(* Logix 5000 project; controller WWTP_CLX vendor 1 type 14 code 54 rev 17.2; software revision 17.00; part 12 of 13 *)
(* tags used below, declared in another part *)
   I_FeedP2_Fault : ALIAS FOR WWTP_CLX_Rack01_Slot00_CNB:I.Slot[1].Data.6;
   I_FeedP2_Fault_IOFault : ALIAS FOR WWTP_CLX_Rack01_Slot00_CNB:I.Slot[1].Fault.6;
   I_FeedP2_InAuto : ALIAS FOR WWTP_CLX_Rack01_Slot00_CNB:I.Slot[1].Data.4;
   I_FeedP2_InAuto_IOFault : ALIAS FOR WWTP_CLX_Rack01_Slot00_CNB:I.Slot[1].Fault.4;
   I_FeedP2_OverLoad : ALIAS FOR WWTP_CLX_Rack01_Slot00_CNB:I.Slot[1].Data.7;
   I_FeedP2_OverLoad_IOFault : ALIAS FOR WWTP_CLX_Rack01_Slot00_CNB:I.Slot[1].Fault.7;
   I_FeedP2_RunFdbk : ALIAS FOR WWTP_CLX_Rack01_Slot00_CNB:I.Slot[1].Data.5;
   I_FeedP2_RunFdbk_IOFault : ALIAS FOR WWTP_CLX_Rack01_Slot00_CNB:I.Slot[1].Fault.5;
   I_FeedP2_SpeedFdbk : ALIAS FOR WWTP_CLX_Rack01_Slot00_CNB:4:I.Ch3Data;
   I_FeedP2_SpeedFdbk_IOFault : ALIAS FOR WWTP_CLX_Rack01_Slot00_CNB:4:I.Ch3Fault;
   O_FeedP2_Out_Run : ALIAS FOR WWTP_CLX_Rack01_Slot00_CNB:2:O.Data.1;
   O_FeedP2_SpeedRef : ALIAS FOR WWTP_CLX_Rack01_Slot00_CNB:6:O.Ch1Data;
   O_FeedP2_SpeedRef_IOFault : ALIAS FOR WWTP_CLX_Rack01_Slot00_CNB:6:I.Ch1Fault;
   PLC_Device_ResetPB : BOOL;   // Site Wide Device Reset Push Button
   PLC_Simulation : BOOL;   // Application running IN SIMULATION
   WWTP_AerTk_InflFlow : UD_Flow;   // Aeration Tank Influent Flow
   WWTP_Alum : UD_Chemical;   // Alum Chemical
   WWTP_AlumTk1Lv : P_AIn;   // Alum Tank #1 Level
   WWTP_FeedP1 : UD_VSD;   // Feed Pump #1
   WWTP_FeedP1_FlowPacing : U_FlowPacing;   // Feed Pump #1 Flow Pacing
   WWTP_FeedP2 : UD_VSD;   // Feed Pump #2
   WWTP_FeedP2_FlowPacing : U_FlowPacing;   // Feed Pump #2 Flow Pacing
   WWTP_FeedP2_OverLoad : P_DIn;   // Feed Pump #2 Overload
   WWTP_FeedSys_OSet_PumpSelect : BOOL;   // Feed Pump System Pump Select
(* FeedP1, continued *)

ROUTINE Main   (* ladder *)
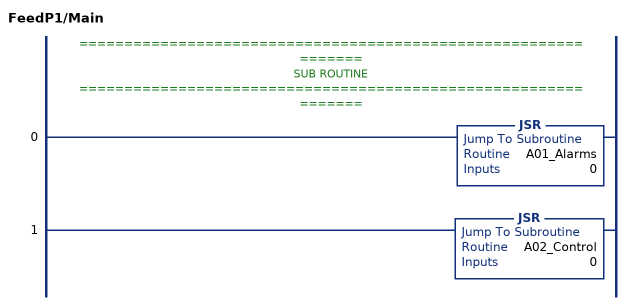
   // ===============================================================
   // SUB ROUTINE
   // ===============================================================
   0: JSR(A01_Alarms,0);
   1: JSR(A02_Control,0);
END_ROUTINE
END_PROGRAM

PROGRAM FeedP2   (* main routine Main *)
VAR
   Device : ALIAS FOR WWTP_FeedP2;
   Device_Alm0 : ALIAS FOR WWTP_FeedP2_OverLoad;
   Device_Alm0_Input : ALIAS FOR I_FeedP2_OverLoad;
   Device_Alm0_Input_IOFault : ALIAS FOR I_FeedP2_OverLoad_IOFault;
   Device_Alm1 : P_DIn := (Inp_Gate := 1, Cfg_NormTextVis := 1, Cfg_PCmdClear := 1, Cfg_TgtDisagreeAckReqd := 1, Cfg_TgtDisagreeSeverity := 3, Sts_InpPV := 1, Ack_TgtDisagree := 1, Rdy_SubstPV := 1);
   Device_Alm1_Input : BOOL;
   Device_Alm1_Input_IOFault : BOOL;
   Device_Alm2 : P_DIn := (Inp_Target := 1, Inp_Gate := 1, Cfg_NormTextVis := 1, Cfg_PCmdClear := 1, Cfg_TgtDisagreeAckReqd := 1, Cfg_TgtDisagreeSeverity := 3, Sts_SubstPV := 1, Sts_TgtDisagree := 1, Ack_TgtDisagree := 1, Rdy_InpPV := 1);
   Device_Alm2_Input : BOOL;
   Device_Alm2_Input_IOFault : BOOL;
   Device_Alm3 : P_DIn := (Inp_Target := 1, Inp_Gate := 1, Cfg_NormTextVis := 1, Cfg_PCmdClear := 1, Cfg_TgtDisagreeAckReqd := 1, Cfg_TgtDisagreeSeverity := 3, Sts_SubstPV := 1, Sts_TgtDisagree := 1, Ack_TgtDisagree := 1, Rdy_InpPV := 1);
   Device_Alm3_Input : BOOL;
   Device_Alm3_Input_IOFault : BOOL;
   Device_Alm4 : P_DIn := (Inp_Target := 1, Inp_Gate := 1, Cfg_NormTextVis := 1, Cfg_PCmdClear := 1, Cfg_TgtDisagreeAckReqd := 1, Cfg_TgtDisagreeSeverity := 3, Sts_SubstPV := 1, Sts_TgtDisagree := 1, Ack_TgtDisagree := 1, Rdy_InpPV := 1);
   Device_Alm4_Input : BOOL;
   Device_Alm4_Input_IOFault : BOOL;
   Device_Faulted : ALIAS FOR I_FeedP2_Fault;
   Device_Faulted_IOFault : ALIAS FOR I_FeedP2_Fault_IOFault;
   Device_GroupReset : ALIAS FOR PLC_Device_ResetPB;
   Device_InAuto : ALIAS FOR I_FeedP2_InAuto;
   Device_InAuto_IOFault : ALIAS FOR I_FeedP2_InAuto_IOFault;
   Device_Out_Run : ALIAS FOR O_FeedP2_Out_Run;
   Device_RunFdbk : ALIAS FOR I_FeedP2_RunFdbk;
   Device_RunFdbk_IOFault : ALIAS FOR I_FeedP2_RunFdbk_IOFault;
   Device_SpeedFdbk : ALIAS FOR I_FeedP2_SpeedFdbk;
   Device_SpeedFdbk_IOFault : ALIAS FOR I_FeedP2_SpeedFdbk_IOFault;
   Device_SpeedRef : ALIAS FOR O_FeedP2_SpeedRef;
   Device_SpeedRef_IOFault : ALIAS FOR O_FeedP2_SpeedRef_IOFault;
END_VAR

ROUTINE A01_Alarms   (* ladder *)
// Discrete Alarms
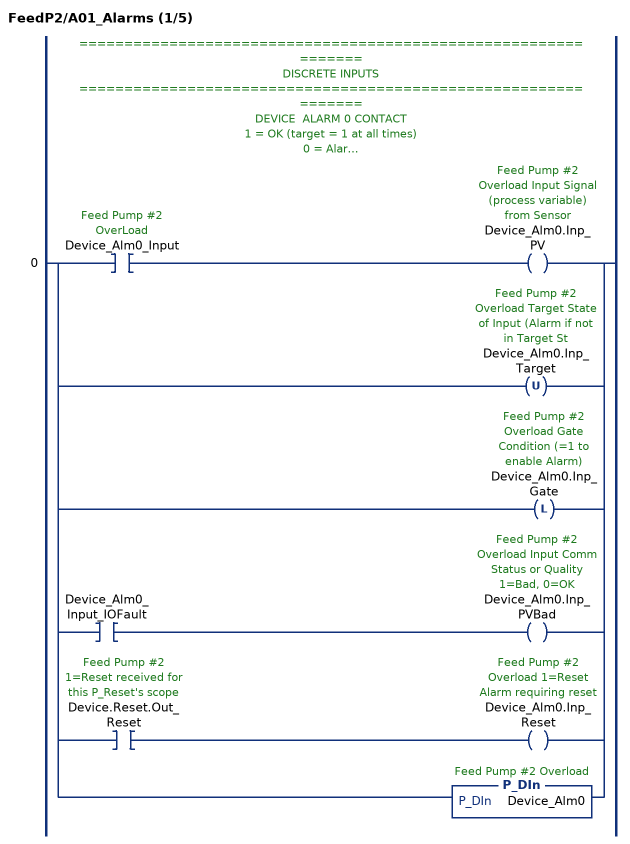
   // ===============================================================
   // DISCRETE INPUTS
   // ===============================================================
   // DEVICE  ALARM 0 CONTACT
   // 1 = OK (target = 1 at all times)
   // 0 = Alarm
   // ALWAYS checked (Gate = 1 at all times)
   0: [XIC(Device_Alm0_Input) OTE(Device_Alm0.Inp_PV) ,OTU(Device_Alm0.Inp_Target) ,OTL(Device_Alm0.Inp_Gate) ,XIC(Device_Alm0_Input_IOFault) OTE(Device_Alm0.Inp_PVBad) ,XIC(Device.Reset.Out_Reset) OTE(Device_Alm0.Inp_Reset) ,P_DIn(Device_Alm0) ];
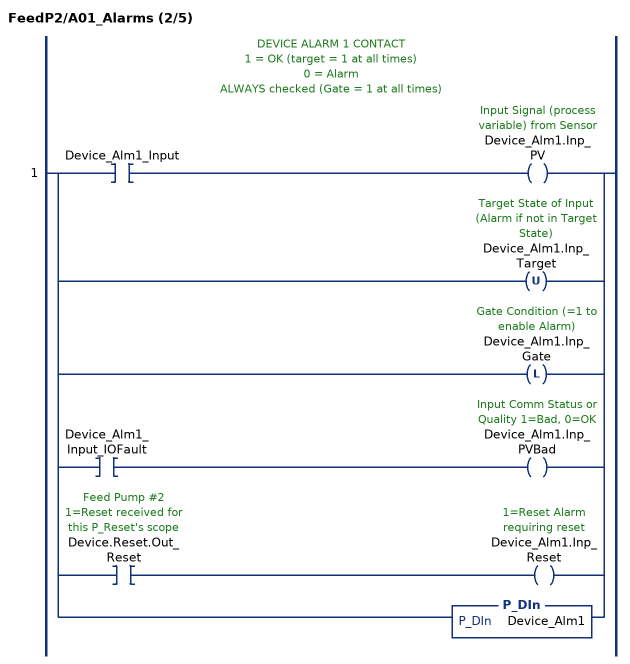
   // DEVICE ALARM 1 CONTACT
   // 1 = OK (target = 1 at all times)
   // 0 = Alarm
   // ALWAYS checked (Gate = 1 at all times)
   1: [XIC(Device_Alm1_Input) OTE(Device_Alm1.Inp_PV) ,OTU(Device_Alm1.Inp_Target) ,OTL(Device_Alm1.Inp_Gate) ,XIC(Device_Alm1_Input_IOFault) OTE(Device_Alm1.Inp_PVBad) ,XIC(Device.Reset.Out_Reset) OTE(Device_Alm1.Inp_Reset) ,P_DIn(Device_Alm1) ];
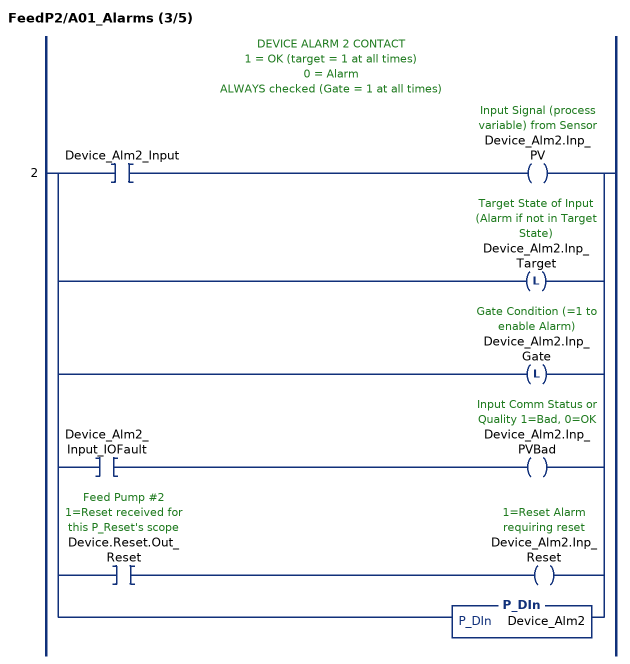
   // DEVICE ALARM 2 CONTACT
   // 1 = OK (target = 1 at all times)
   // 0 = Alarm
   // ALWAYS checked (Gate = 1 at all times)
   2: [XIC(Device_Alm2_Input) OTE(Device_Alm2.Inp_PV) ,OTL(Device_Alm2.Inp_Target) ,OTL(Device_Alm2.Inp_Gate) ,XIC(Device_Alm2_Input_IOFault) OTE(Device_Alm2.Inp_PVBad) ,XIC(Device.Reset.Out_Reset) OTE(Device_Alm2.Inp_Reset) ,P_DIn(Device_Alm2) ];
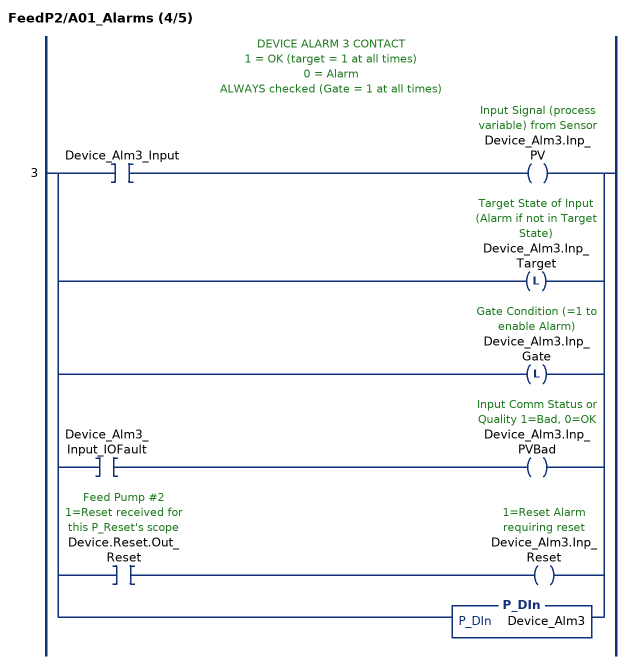
   // DEVICE ALARM 3 CONTACT
   // 1 = OK (target = 1 at all times)
   // 0 = Alarm
   // ALWAYS checked (Gate = 1 at all times)
   3: [XIC(Device_Alm3_Input) OTE(Device_Alm3.Inp_PV) ,OTL(Device_Alm3.Inp_Target) ,OTL(Device_Alm3.Inp_Gate) ,XIC(Device_Alm3_Input_IOFault) OTE(Device_Alm3.Inp_PVBad) ,XIC(Device.Reset.Out_Reset) OTE(Device_Alm3.Inp_Reset) ,P_DIn(Device_Alm3) ];
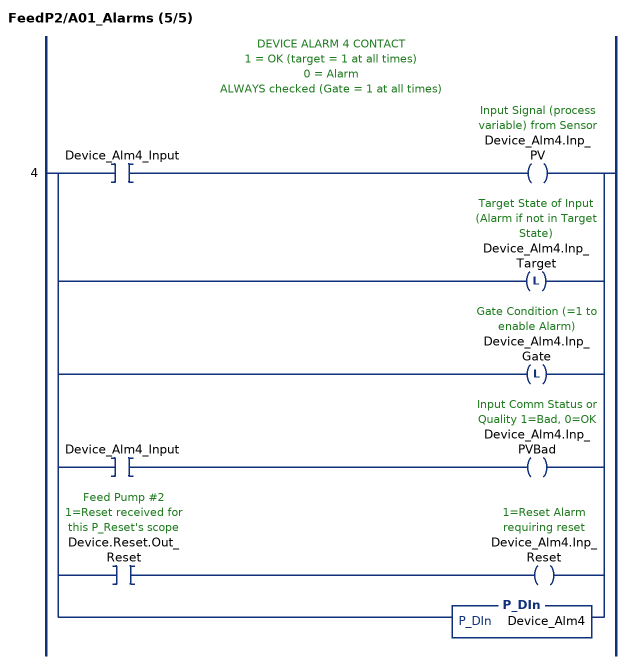
   // DEVICE ALARM 4 CONTACT
   // 1 = OK (target = 1 at all times)
   // 0 = Alarm
   // ALWAYS checked (Gate = 1 at all times)
   4: [XIC(Device_Alm4_Input) OTE(Device_Alm4.Inp_PV) ,OTL(Device_Alm4.Inp_Target) ,OTL(Device_Alm4.Inp_Gate) ,XIC(Device_Alm4_Input) OTE(Device_Alm4.Inp_PVBad) ,XIC(Device.Reset.Out_Reset) OTE(Device_Alm4.Inp_Reset) ,P_DIn(Device_Alm4) ];
END_ROUTINE

ROUTINE A02_Control   (* ladder *)
// Device Contol
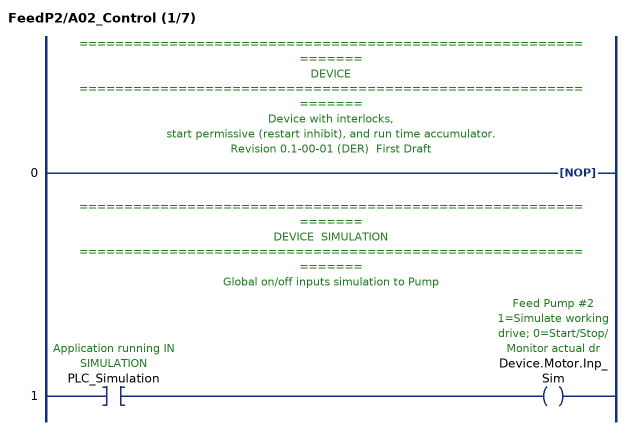
   // ===============================================================
   // DEVICE
   // ===============================================================
   // Device with interlocks,
   // start permissive (restart inhibit), and run time accumulator.
   // Revision 0.1-00-01 (DER)  First Draft
   0: NOP();
   // ===============================================================
   // DEVICE  SIMULATION
   // ===============================================================
   // Global on/off inputs simulation to Pump
   1: XIC(PLC_Simulation)OTE(Device.Motor.Inp_Sim);
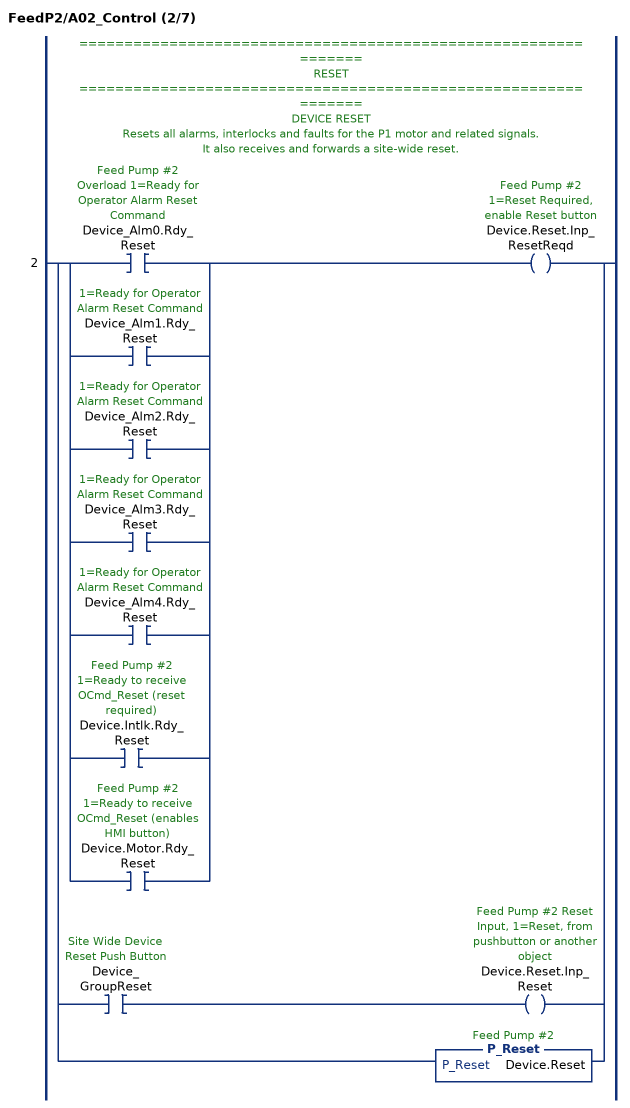
   // ===============================================================
   // RESET
   // ===============================================================
   // DEVICE RESET
   // Resets all alarms, interlocks and faults for the P1 motor and related signals.
   // It also receives and forwards a site-wide reset.
   2: [[XIC(Device_Alm0.Rdy_Reset) ,XIC(Device_Alm1.Rdy_Reset) ,XIC(Device_Alm2.Rdy_Reset) ,XIC(Device_Alm3.Rdy_Reset) ,XIC(Device_Alm4.Rdy_Reset) ,XIC(Device.Intlk.Rdy_Reset) ,XIC(Device.Motor.Rdy_Reset) ] OTE(Device.Reset.Inp_ResetReqd) ,XIC(Device_GroupReset) OTE(Device.Reset.Inp_Reset) ,P_Reset(Device.Reset) ];
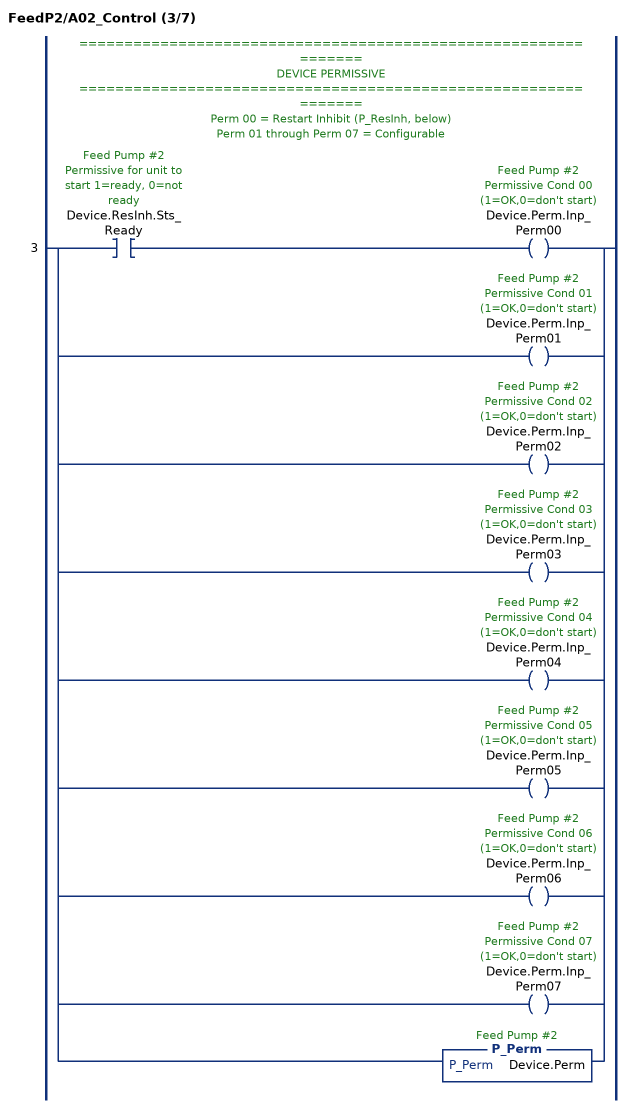
   // ===============================================================
   // DEVICE PERMISSIVE
   // ===============================================================
   // Perm 00 = Restart Inhibit (P_ResInh, below)
   // Perm 01 through Perm 07 = Configurable
   3: [XIC(Device.ResInh.Sts_Ready) OTE(Device.Perm.Inp_Perm00) ,OTE(Device.Perm.Inp_Perm01) ,OTE(Device.Perm.Inp_Perm02) ,OTE(Device.Perm.Inp_Perm03) ,OTE(Device.Perm.Inp_Perm04) ,OTE(Device.Perm.Inp_Perm05) ,OTE(Device.Perm.Inp_Perm06) ,OTE(Device.Perm.Inp_Perm07) ,P_Perm(Device.Perm) ];
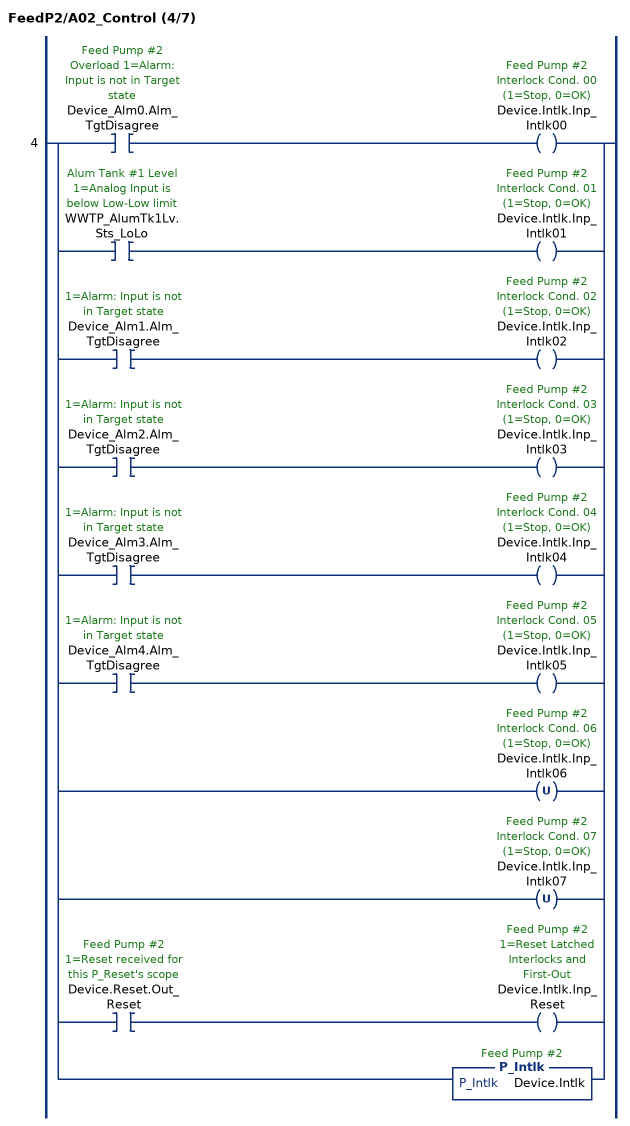
   4: [XIC(Device_Alm0.Alm_TgtDisagree) OTE(Device.Intlk.Inp_Intlk00) ,XIC(WWTP_AlumTk1Lv.Sts_LoLo) OTE(Device.Intlk.Inp_Intlk01) ,XIC(Device_Alm1.Alm_TgtDisagree) OTE(Device.Intlk.Inp_Intlk02) ,XIC(Device_Alm2.Alm_TgtDisagree) OTE(Device.Intlk.Inp_Intlk03) ,XIC(Device_Alm3.Alm_TgtDisagree) OTE(Device.Intlk.Inp_Intlk04) ,XIC(Device_Alm4.Alm_TgtDisagree) OTE(Device.Intlk.Inp_Intlk05) ,OTU(Device.Intlk.Inp_Intlk06) ,OTU(Device.Intlk.Inp_Intlk07) ,XIC(Device.Reset.Out_Reset) OTE(Device.Intlk.Inp_Reset) ,P_Intlk(Device.Intlk) ];
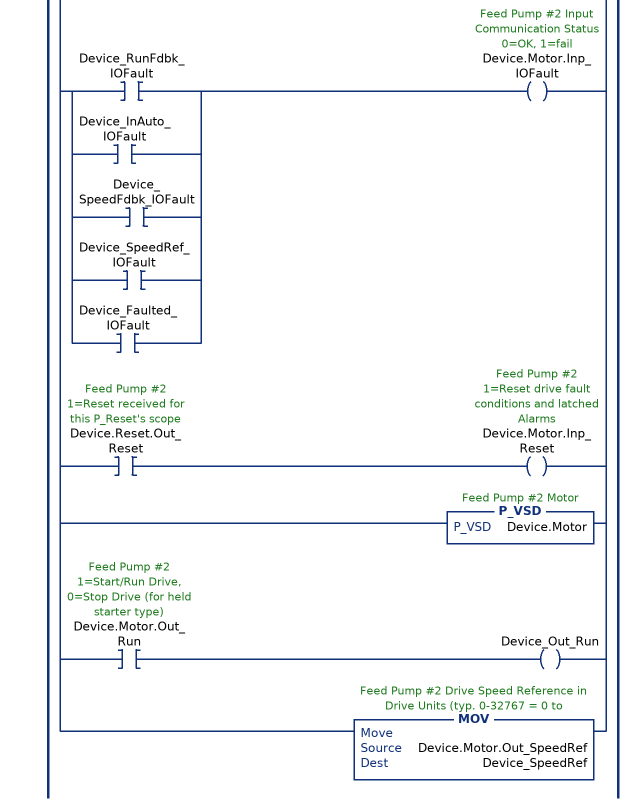
   // ===============================================================
   // DEVICE MOTOR
   // ===============================================================
   // This rung actually monitors and controls the Device motor.
   // Mapping inputs:  Run Feedback
   // Hand Mode selection (local operation)
   // Permissive OK
   // Protective’s OK,
   // I/O Fault signals
   // Pump Reset (above)
   // DEVICE
   // Output Mapping: Starter output
   5: [XIC(Device_RunFdbk) OTE(Device.Motor.Inp_Running) ,MOV(Device_SpeedFdbk,Device.Motor.Inp_SpeedFdbk) ,XIO(Device_InAuto) OTE(Device.Motor.Inp_Hand) ,XIC(Device_Faulted) OTE(Device.Motor.Inp_Faulted) ,XIC(Device.Perm.Sts_PermOK) OTE(Device.Motor.Inp_FwdPermOK) ,XIC(Device.Perm.Sts_NBPermOK) OTE(Device.Motor.Inp_FwdNBPermOK) ,XIC(Device.Intlk.Sts_IntlkOK) OTE(Device.Motor.Inp_IntlkOK) ,XIC(Device.Intlk.Sts_NBIntlkOK) OTE(Device.Motor.Inp_NBIntlkOK) ,[XIC(Device_RunFdbk_IOFault) ,XIC(Device_InAuto_IOFault) ,XIC(Device_SpeedFdbk_IOFault) ,XIC(Device_SpeedRef_IOFault) ,XIC(Device_Faulted_IOFault) ] OTE(Device.Motor.Inp_IOFault) ,XIC(Device.Reset.Out_Reset) OTE(Device.Motor.Inp_Reset) ,P_VSD(Device.Motor) ,XIC(Device.Motor.Out_Run) OTE(Device_Out_Run) ,MOV(Device.Motor.Out_SpeedRef,Device_SpeedRef) ];
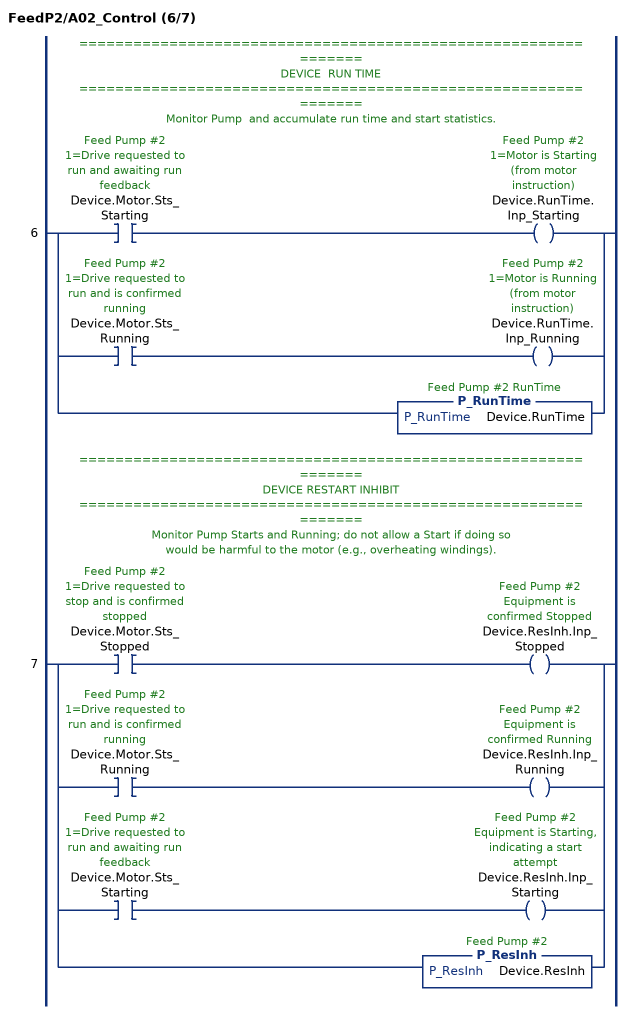
   // ===============================================================
   // DEVICE  RUN TIME
   // ===============================================================
   // Monitor Pump  and accumulate run time and start statistics.
   6: [XIC(Device.Motor.Sts_Starting) OTE(Device.RunTime.Inp_Starting) ,XIC(Device.Motor.Sts_Running) OTE(Device.RunTime.Inp_Running) ,P_RunTime(Device.RunTime) ];
   // ===============================================================
   // DEVICE RESTART INHIBIT
   // ===============================================================
   // Monitor Pump Starts and Running; do not allow a Start if doing so
   // would be harmful to the motor (e.g., overheating windings).
   7: [XIC(Device.Motor.Sts_Stopped) OTE(Device.ResInh.Inp_Stopped) ,XIC(Device.Motor.Sts_Running) OTE(Device.ResInh.Inp_Running) ,XIC(Device.Motor.Sts_Starting) OTE(Device.ResInh.Inp_Starting) ,P_ResInh(Device.ResInh) ];
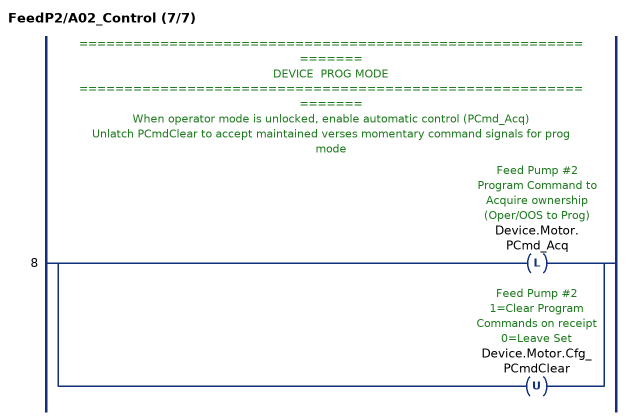
   // ===============================================================
   // DEVICE  PROG MODE
   // ===============================================================
   // When operator mode is unlocked, enable automatic control (PCmd_Acq)
   // Unlatch PCmdClear to accept maintained verses momentary command signals for prog mode
   8: [OTL(Device.Motor.PCmd_Acq) ,OTU(Device.Motor.Cfg_PCmdClear) ];
END_ROUTINE

ROUTINE Main   (* ladder *)
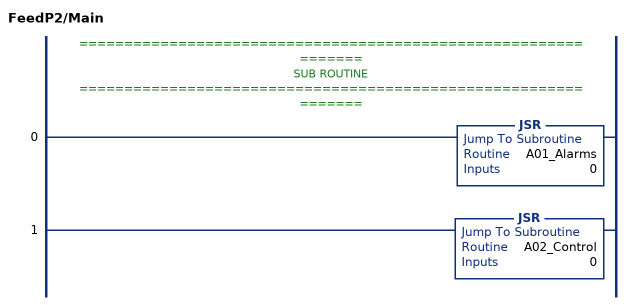
   // ===============================================================
   // SUB ROUTINE
   // ===============================================================
   0: JSR(A01_Alarms,0);
   1: JSR(A02_Control,0);
END_ROUTINE
END_PROGRAM

PROGRAM FeedPSys   (* main routine Main *)
VAR
   Chemical : ALIAS FOR WWTP_Alum;
   P1_FlowPacing : ALIAS FOR WWTP_FeedP1_FlowPacing;
   P1_Motor : ALIAS FOR WWTP_FeedP1.Motor;
   P2_FlowPacing : ALIAS FOR WWTP_FeedP2_FlowPacing;
   P2_Motor : ALIAS FOR WWTP_FeedP2.Motor;
   PacedFlow : ALIAS FOR WWTP_AerTk_InflFlow;
   PumpSelect : ALIAS FOR WWTP_FeedSys_OSet_PumpSelect;
END_VAR

ROUTINE A01_Control   (* ladder *)
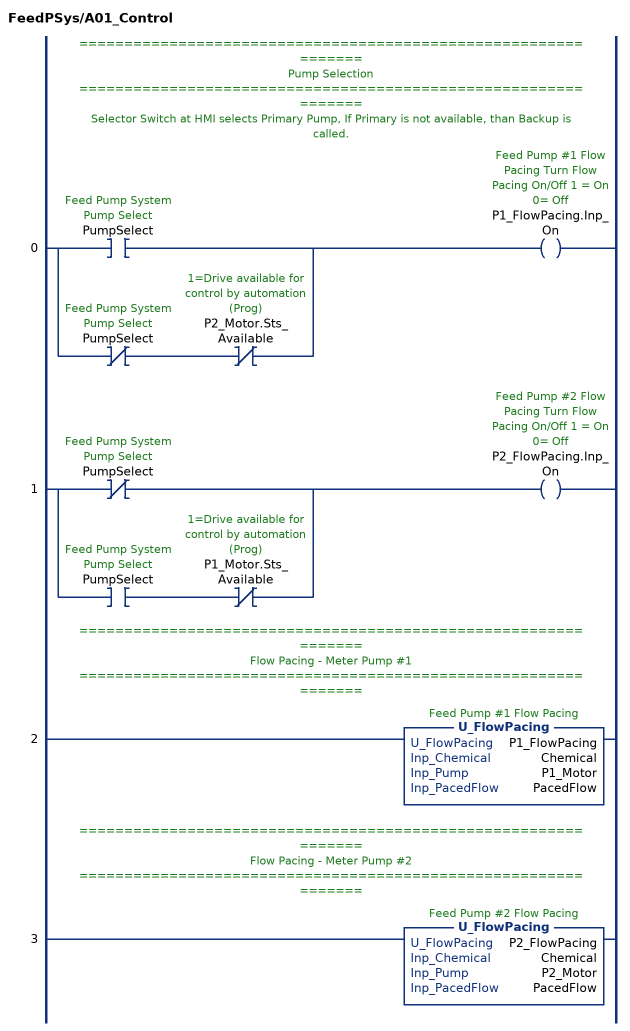
   // ===============================================================
   // Pump Selection
   // ===============================================================
   // Selector Switch at HMI selects Primary Pump, If Primary is not available, than Backup is called.
   0: [XIC(PumpSelect) ,XIO(PumpSelect) XIO(P2_Motor.Sts_Available) ]OTE(P1_FlowPacing.Inp_On);
   1: [XIO(PumpSelect) ,XIC(PumpSelect) XIO(P1_Motor.Sts_Available) ]OTE(P2_FlowPacing.Inp_On);
   // ===============================================================
   // Flow Pacing - Meter Pump #1
   // ===============================================================
   2: U_FlowPacing(P1_FlowPacing,Chemical,P1_Motor,PacedFlow);
   // ===============================================================
   // Flow Pacing - Meter Pump #2
   // ===============================================================
   3: U_FlowPacing(P2_FlowPacing,Chemical,P2_Motor,PacedFlow);
END_ROUTINE

ROUTINE Main   (* ladder *)
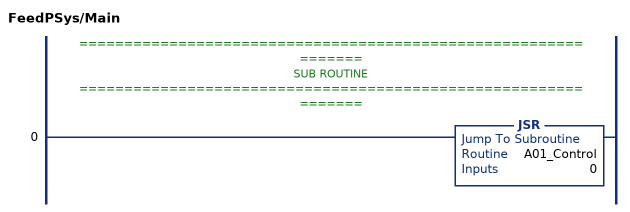
   // ===============================================================
   // SUB ROUTINE
   // ===============================================================
   0: JSR(A01_Control,0);
END_ROUTINE
END_PROGRAM

PROGRAM MainProgram   (* main routine Main *)
VAR
   Alm00 : P_DIn := (Inp_Target := 1, Inp_Gate := 1, Inp_Reset := 1, Cfg_NormTextVis := 1, Cfg_PCmdClear := 1, Cfg_TgtDisagreeAckReqd := 1, Cfg_TgtDisagreeSeverity := 3, Sts_InpPV := 1, Sts_TgtDisagree := 1, Ack_TgtDisagree := 1, Rdy_SubstPV := 1);
   Alm00_Input : BOOL;
   Alm00_Input_IOFault : BOOL;
   Alm01 : P_DIn := (Inp_Target := 1, Inp_Gate := 1, Inp_Reset := 1, Cfg_NormTextVis := 1, Cfg_PCmdClear := 1, Cfg_TgtDisagreeAckReqd := 1, Cfg_TgtDisagreeSeverity := 3, Sts_InpPV := 1, Sts_TgtDisagree := 1, Ack_TgtDisagree := 1, Rdy_SubstPV := 1);
   Alm01_Input : BOOL;
   Alm01_Input_IOFault : BOOL;
   Alm02 : P_DIn := (Inp_Target := 1, Inp_Gate := 1, Inp_Reset := 1, Cfg_NormTextVis := 1, Cfg_PCmdClear := 1, Cfg_TgtDisagreeAckReqd := 1, Cfg_TgtDisagreeSeverity := 3, Sts_SubstPV := 1, Sts_TgtDisagree := 1, Ack_TgtDisagree := 1, Rdy_InpPV := 1);
   Alm02_Input : BOOL;
   Alm02_Input_IOFault : BOOL;
   Alm03 : P_DIn := (Inp_Target := 1, Inp_Gate := 1, Inp_Reset := 1, Cfg_NormTextVis := 1, Cfg_PCmdClear := 1, Cfg_TgtDisagreeAckReqd := 1, Cfg_TgtDisagreeSeverity := 3, Sts_SubstPV := 1, Sts_TgtDisagree := 1, Ack_TgtDisagree := 1, Rdy_InpPV := 1);
   Alm03_Input : BOOL;
   Alm03_Input_IOFault : BOOL;
   Alm04 : P_DIn := (Inp_Target := 1, Inp_Gate := 1, Inp_Reset := 1, Cfg_NormTextVis := 1, Cfg_PCmdClear := 1, Cfg_TgtDisagreeAckReqd := 1, Cfg_TgtDisagreeSeverity := 3, Sts_SubstPV := 1, Sts_TgtDisagree := 1, Ack_TgtDisagree := 1, Rdy_InpPV := 1);
   Alm04_Input : BOOL;
   Alm04_Input_IOFault : BOOL;
END_VAR

ROUTINE A01_DiscreteInputs   (* ladder *)
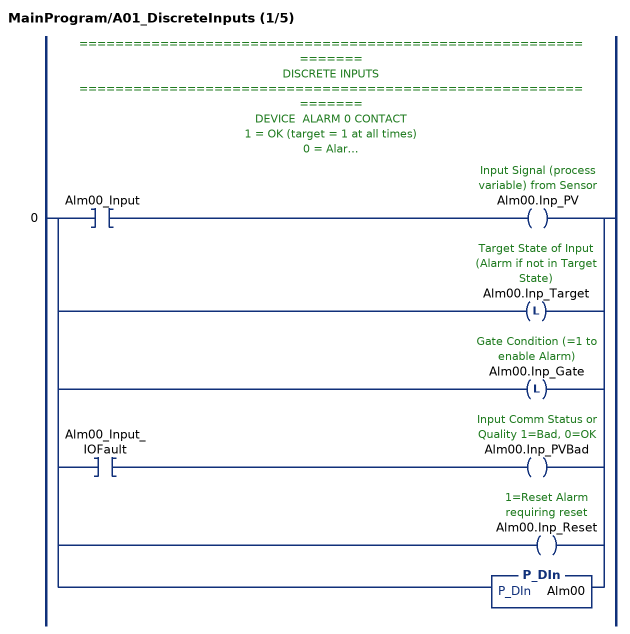
   // ===============================================================
   // DISCRETE INPUTS
   // ===============================================================
   // DEVICE  ALARM 0 CONTACT
   // 1 = OK (target = 1 at all times)
   // 0 = Alarm
   // ALWAYS checked (Gate = 1 at all times)
   0: [XIC(Alm00_Input) OTE(Alm00.Inp_PV) ,OTL(Alm00.Inp_Target) ,OTL(Alm00.Inp_Gate) ,XIC(Alm00_Input_IOFault) OTE(Alm00.Inp_PVBad) ,OTE(Alm00.Inp_Reset) ,P_DIn(Alm00) ];
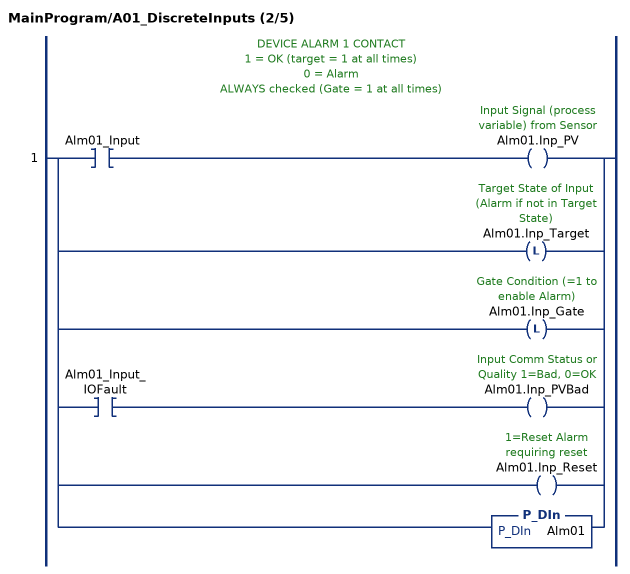
   // DEVICE ALARM 1 CONTACT
   // 1 = OK (target = 1 at all times)
   // 0 = Alarm
   // ALWAYS checked (Gate = 1 at all times)
   1: [XIC(Alm01_Input) OTE(Alm01.Inp_PV) ,OTL(Alm01.Inp_Target) ,OTL(Alm01.Inp_Gate) ,XIC(Alm01_Input_IOFault) OTE(Alm01.Inp_PVBad) ,OTE(Alm01.Inp_Reset) ,P_DIn(Alm01) ];
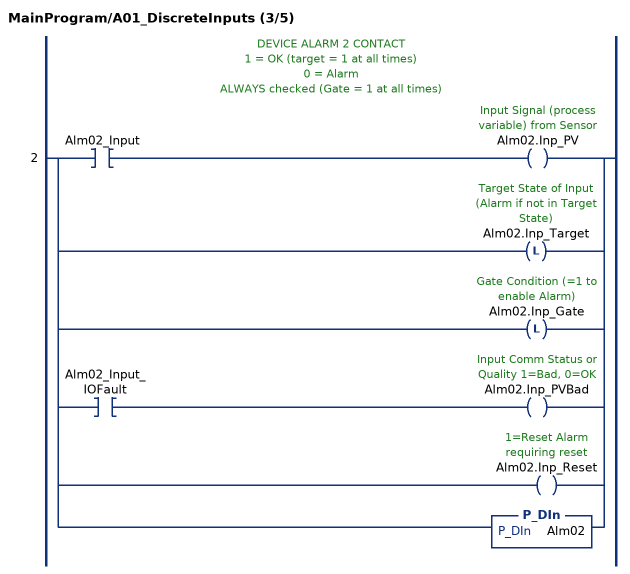
   // DEVICE ALARM 2 CONTACT
   // 1 = OK (target = 1 at all times)
   // 0 = Alarm
   // ALWAYS checked (Gate = 1 at all times)
   2: [XIC(Alm02_Input) OTE(Alm02.Inp_PV) ,OTL(Alm02.Inp_Target) ,OTL(Alm02.Inp_Gate) ,XIC(Alm02_Input_IOFault) OTE(Alm02.Inp_PVBad) ,OTE(Alm02.Inp_Reset) ,P_DIn(Alm02) ];
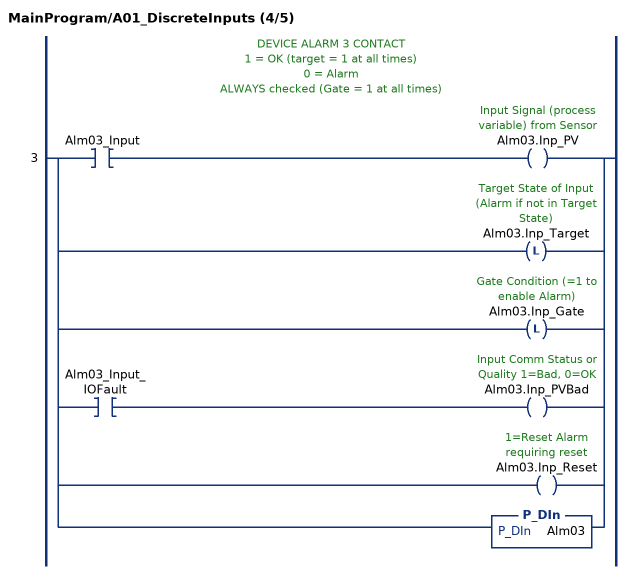
   // DEVICE ALARM 3 CONTACT
   // 1 = OK (target = 1 at all times)
   // 0 = Alarm
   // ALWAYS checked (Gate = 1 at all times)
   3: [XIC(Alm03_Input) OTE(Alm03.Inp_PV) ,OTL(Alm03.Inp_Target) ,OTL(Alm03.Inp_Gate) ,XIC(Alm03_Input_IOFault) OTE(Alm03.Inp_PVBad) ,OTE(Alm03.Inp_Reset) ,P_DIn(Alm03) ];
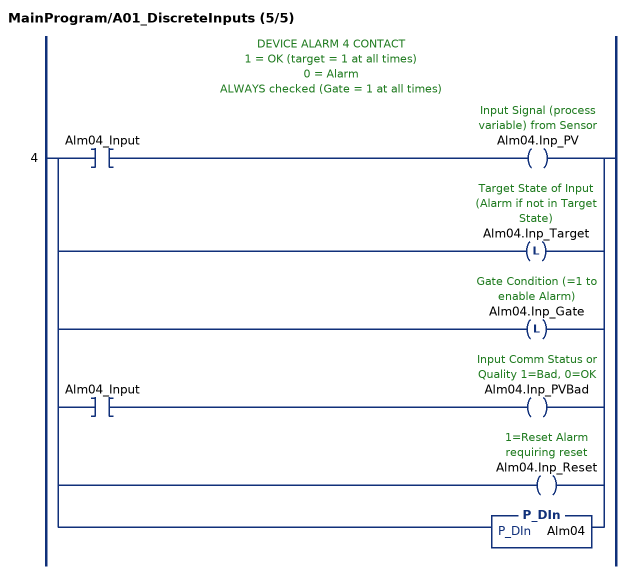
   // DEVICE ALARM 4 CONTACT
   // 1 = OK (target = 1 at all times)
   // 0 = Alarm
   // ALWAYS checked (Gate = 1 at all times)
   4: [XIC(Alm04_Input) OTE(Alm04.Inp_PV) ,OTL(Alm04.Inp_Target) ,OTL(Alm04.Inp_Gate) ,XIC(Alm04_Input) OTE(Alm04.Inp_PVBad) ,OTE(Alm04.Inp_Reset) ,P_DIn(Alm04) ];
END_ROUTINE
